RoboDK station: Bench V1 cell v7.rdk

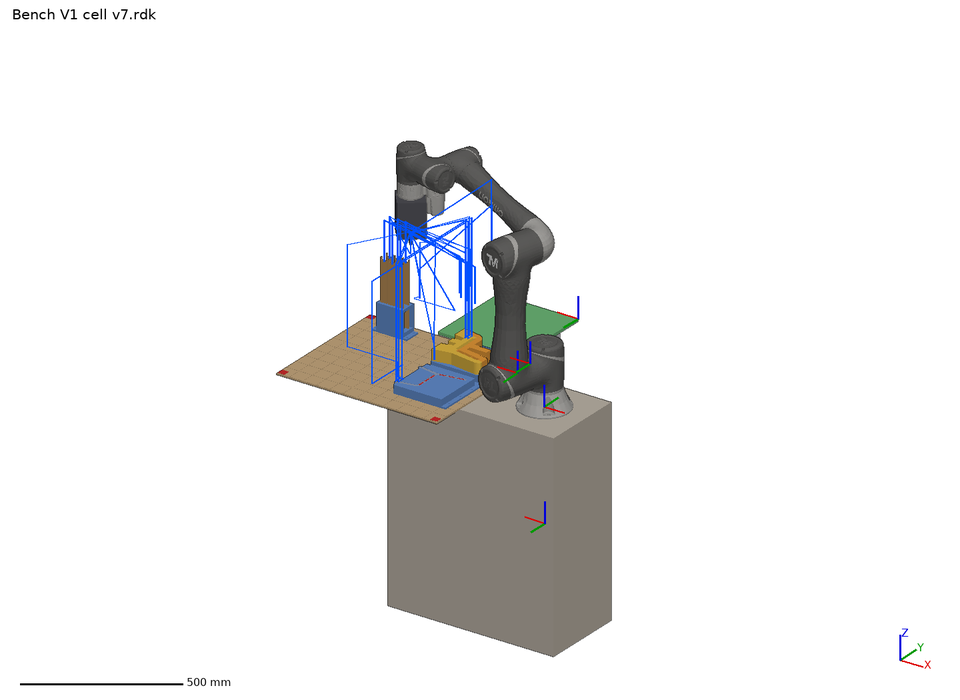
[picture v0: the station drawn from its stored meshes, robots at their saved joint values, targets as dots, program paths as lines]
Station Bench V1 cell v7 (saved by RoboDK 6.1.1). Poses are relative to the parent item; angles as X-Y-Z fixed-axis rotations.
  - frame Cell at (0, 0, 0) mm
    - frame Work plate at (-206.44, 152.99, -4.46) mm, rotated rx -0.03 ry -0.07 rz -179.98 deg
      - frame Ground base at (0, -67, 6) mm
        - object Table at (0, 0, 0) mm, size 620 x 310 x 744 mm
        - object Ground base plate at (0, 0, 0) mm, size 600 x 500 x 6 mm, geometry from ground_base_v7.stl
        - object Vision square 1 at (3, 3, 0) mm, size 25 x 25 x 0.5 mm, geometry from vision_square.stl
        - object Vision square 2 at (3, 472, 0) mm, size 25 x 25 x 0.5 mm, geometry from vision_square.stl
        - object Vision square 3 at (572, 3, 0) mm, size 25 x 25 x 0.5 mm, geometry from vision_square.stl
        - object Vision square 4 at (572, 472, 0) mm, size 25 x 25 x 0.5 mm, geometry from vision_square.stl
        - object Base A at (135, 122, 10) mm, rotated rx 0 ry 0 rz 90 deg, size 196 x 196 x 30 mm, geometry from base_a_v7.stl
        - object Base B at (135, 322, 10) mm, rotated rx 0 ry 0 rz -90 deg, size 196 x 196 x 30 mm, geometry from base_b_v7.stl
        - object Plank jig at (420, 30, 0) mm, size 132 x 60 x 100 mm, geometry from plank_rack_v7.stl
        - frame AMR at (60, -340, 0) mm
          - object AMR plate at (0, 0, 0) mm, size 300 x 320 x 10 mm
          - object AMR top module at (0, 0, 0) mm, size 220 x 240 x 363 mm
          - frame Omron LD-250 Base at (150, -40, -756) mm
            - robot AMR LD-250: 4 axes
                joint limits [-10000, -10000, -10, -3600] to [10000, 10000, 10, 3600]; home [0, 0, 0, 0]; saved at [0, 0, 0, 0]
        - object frame1 at (161.88, 119.28, 144.5) mm, size 174.7 x 141.9 x 10 mm, geometry from frame.stl
        - object frame2 at (161.88, 324.71, -95.5) mm, rotated rx 180 ry 0 rz 0 deg, size 174.7 x 141.9 x 10 mm, geometry from frame.stl
        - object piece A1 at (156.88, 119.28, 144.5) mm, rotated rx 90 ry 0 rz 90 deg, size 21.4 x 10 x 5 mm, geometry from interface_piece.stl
        - object piece B1 at (156.88, 324.71, 144.5) mm, rotated rx 90 ry 0 rz 90 deg, size 21.4 x 10 x 5 mm, geometry from interface_piece.stl
        - object plank1 at (435, 47.5, 128) mm, rotated rx 90 ry 0 rz 0 deg, size 25 x 250 x 5 mm, geometry from plank_body.stl
        - object piece A2 at (156.88, 89.3, 144.5) mm, rotated rx 90 ry 0 rz 90 deg, size 21.4 x 10 x 5 mm, geometry from interface_piece.stl
        - object piece B2 at (156.88, 354.7, 144.5) mm, rotated rx 90 ry 0 rz 90 deg, size 21.4 x 10 x 5 mm, geometry from interface_piece.stl
        - object plank2 at (465, 47.5, 128) mm, rotated rx 90 ry 0 rz 0 deg, size 25 x 250 x 5 mm, geometry from plank_body.stl
        - object piece A3 at (156.88, 149.27, 144.5) mm, rotated rx 90 ry 0 rz 90 deg, size 21.4 x 10 x 5 mm, geometry from interface_piece.stl
        - object piece B3 at (156.88, 294.73, 144.5) mm, rotated rx 90 ry 0 rz 90 deg, size 21.4 x 10 x 5 mm, geometry from interface_piece.stl
        - object plank3 at (495, 47.5, 128) mm, rotated rx 90 ry 0 rz 0 deg, size 25 x 250 x 5 mm, geometry from plank_body.stl
        - object piece A4 at (138.44, 171.24, 144.5) mm, rotated rx 90 ry 0 rz 170 deg, size 21.4 x 10 x 5 mm, geometry from interface_piece.stl
        - object piece B4 at (138.44, 272.76, 144.5) mm, rotated rx 90 ry 0 rz 10 deg, size 21.4 x 10 x 5 mm, geometry from interface_piece.stl
        - object plank4 at (435, 77.5, 128) mm, rotated rx 90 ry 0 rz 0 deg, size 25 x 250 x 5 mm, geometry from plank_body.stl
        - object piece A5 at (108.91, 176.45, 144.5) mm, rotated rx 90 ry 0 rz 170 deg, size 21.4 x 10 x 5 mm, geometry from interface_piece.stl
        - object piece B5 at (108.91, 267.55, 144.5) mm, rotated rx 90 ry 0 rz 10 deg, size 21.4 x 10 x 5 mm, geometry from interface_piece.stl
        - object plank5 at (465, 77.5, 128) mm, rotated rx 90 ry 0 rz 0 deg, size 25 x 250 x 5 mm, geometry from plank_body.stl
        - object piece A6 at (79.38, 181.66, 144.5) mm, rotated rx 90 ry 0 rz 170 deg, size 21.4 x 10 x 5 mm, geometry from interface_piece.stl
        - object piece B6 at (79.38, 262.34, 144.5) mm, rotated rx 90 ry 0 rz 10 deg, size 21.4 x 10 x 5 mm, geometry from interface_piece.stl
        - object plank6 at (495, 77.5, 128) mm, rotated rx 90 ry 0 rz 0 deg, size 25 x 250 x 5 mm, geometry from plank_body.stl
        - object Guide inner at (135, 122, 10) mm, rotated rx 0 ry 0 rz 90 deg, size 158.3 x 160 x 40 mm, geometry from guide_inner_v7.stl
        - object Guide outer at (135, 122, 10) mm, rotated rx 0 ry 0 rz 90 deg, size 177.7 x 180 x 40 mm, geometry from guide_outer_v7.stl
        - target Home (Cartesian target) at (295, 220, 380) mm, rotated rx 180 ry 0 rz 0 deg; joints [-14.089, 3.172, -81.623, -11.478, -90.01, 75.887] of Omron TM5-900
        - target plank3 pick travel (Cartesian target) at (495, 45, 380) mm, rotated rx 180 ry 0 rz -90 deg; joints [-23.734, -30.79, -38.937, -20.201, -89.998, 156.242] of Omron TM5-900
        - target plank3 pick approach (Cartesian target) at (495, 45, 278) mm, rotated rx 180 ry 0 rz -90 deg; joints [-23.733, -27.058, -59.189, -3.681, -89.998, 156.243] of Omron TM5-900
        - target plank3 pick (Cartesian target) at (495, 45, 238) mm, rotated rx 180 ry 0 rz -90 deg; joints [-23.733, -26.967, -64.904, 1.942, -89.998, 156.243] of Omron TM5-900
        - target plank3 pick out (Cartesian target) at (495, 45, 298) mm, rotated rx 180 ry 0 rz -90 deg; joints [-23.733, -27.342, -55.969, -6.617, -89.998, 156.243] of Omron TM5-900
        - target plank3 pick up (Cartesian target) at (495, 45, 380) mm, rotated rx 180 ry 0 rz -90 deg; joints [-23.734, -30.79, -38.937, -20.201, -89.998, 156.242] of Omron TM5-900
        - target plank3 place travel (Cartesian target) at (159.38, 149.27, 380) mm, rotated rx 180 ry 0 rz 0 deg; joints [-30.116, 20.707, -95.296, -15.34, -89.99, 59.86] of Omron TM5-900
        - target plank3 above guide (Cartesian target) at (159.38, 149.27, 329.5) mm, rotated rx 180 ry 0 rz 0 deg; joints [-30.114, 22.129, -103.368, -8.691, -89.99, 59.862] of Omron TM5-900
        - target plank3 place (Cartesian target) at (159.38, 149.27, 254.5) mm, rotated rx 180 ry 0 rz 0 deg; joints [-30.112, 22.789, -114.254, 1.536, -89.99, 59.864] of Omron TM5-900
        - target plank3 push approach (Cartesian target) at (159.38, 149.27, 289.5) mm, rotated rx 180 ry 0 rz 0 deg; joints [-30.113, 22.711, -109.326, -3.314, -89.99, 59.863] of Omron TM5-900
        - target plank3 push (Cartesian target) at (159.38, 149.27, 269.5) mm, rotated rx 180 ry 0 rz 0 deg; joints [-30.113, 22.808, -112.174, -0.563, -89.99, 59.863] of Omron TM5-900
        - target plank3 push out (Cartesian target) at (159.38, 149.27, 289.5) mm, rotated rx 180 ry 0 rz 0 deg; joints [-30.113, 22.711, -109.326, -3.314, -89.99, 59.863] of Omron TM5-900
        - target plank3 place up (Cartesian target) at (159.38, 149.27, 380) mm, rotated rx 180 ry 0 rz 0 deg; joints [-30.116, 20.707, -95.296, -15.34, -89.99, 59.86] of Omron TM5-900
        - target plank6 pick travel (Cartesian target) at (495, 75, 380) mm, rotated rx 180 ry 0 rz -90 deg; joints [-21.493, -29.466, -41.001, -19.462, -90.001, 158.482] of Omron TM5-900
        - target plank6 pick approach (Cartesian target) at (495, 75, 278) mm, rotated rx 180 ry 0 rz -90 deg; joints [-21.494, -26.016, -60.721, -3.192, -90.001, 158.482] of Omron TM5-900
        - target plank6 pick (Cartesian target) at (495, 75, 238) mm, rotated rx 180 ry 0 rz -90 deg; joints [-21.494, -25.975, -66.359, 2.406, -90.001, 158.482] of Omron TM5-900
        - target plank6 pick out (Cartesian target) at (495, 75, 298) mm, rotated rx 180 ry 0 rz -90 deg; joints [-21.494, -26.268, -57.554, -6.106, -90.001, 158.482] of Omron TM5-900
        - target plank6 pick up (Cartesian target) at (495, 75, 380) mm, rotated rx 180 ry 0 rz -90 deg; joints [-21.493, -29.466, -41.001, -19.462, -90.001, 158.482] of Omron TM5-900
        - target plank6 place travel (Cartesian target) at (79.82, 184.12, 380) mm, rotated rx 180 ry 0 rz 80 deg; joints [-32.257, 32.355, -101.249, -21.035, -89.987, -22.281] of Omron TM5-900
        - target plank6 above guide (Cartesian target) at (79.82, 184.12, 329.5) mm, rotated rx 180 ry 0 rz 80 deg; joints [-32.254, 34.514, -109.51, -14.934, -89.987, -22.278] of Omron TM5-900
        - target plank6 place (Cartesian target) at (79.82, 184.12, 254.5) mm, rotated rx 180 ry 0 rz 80 deg; joints [-32.25, 36.477, -120.901, -5.506, -89.987, -22.275] of Omron TM5-900
        - target plank6 push approach (Cartesian target) at (79.82, 184.12, 289.5) mm, rotated rx 180 ry 0 rz 80 deg; joints [-32.252, 35.762, -115.703, -9.988, -89.987, -22.276] of Omron TM5-900
        - target plank6 push (Cartesian target) at (79.82, 184.12, 269.5) mm, rotated rx 180 ry 0 rz 80 deg; joints [-32.251, 36.217, -118.697, -7.449, -89.987, -22.275] of Omron TM5-900
        - target plank6 push out (Cartesian target) at (79.82, 184.12, 289.5) mm, rotated rx 180 ry 0 rz 80 deg; joints [-32.252, 35.762, -115.703, -9.988, -89.987, -22.276] of Omron TM5-900
        - target plank6 place up (Cartesian target) at (79.82, 184.12, 380) mm, rotated rx 180 ry 0 rz 80 deg; joints [-32.257, 32.355, -101.249, -21.035, -89.987, -22.281] of Omron TM5-900
        - target plank2 pick travel (Cartesian target) at (465, 45, 380) mm, rotated rx 180 ry 0 rz -90 deg; joints [-24.747, -25.325, -47.241, -17.362, -89.997, 155.229] of Omron TM5-900
        - target plank2 pick approach (Cartesian target) at (465, 45, 278) mm, rotated rx 180 ry 0 rz -90 deg; joints [-24.747, -22.614, -65.589, -1.725, -89.997, 155.229] of Omron TM5-900
        - target plank2 pick (Cartesian target) at (465, 45, 238) mm, rotated rx 180 ry 0 rz -90 deg; joints [-24.746, -22.719, -71.021, 3.812, -89.997, 155.229] of Omron TM5-900
        - target plank2 pick out (Cartesian target) at (465, 45, 298) mm, rotated rx 180 ry 0 rz -90 deg; joints [-24.747, -22.777, -62.567, -4.584, -89.997, 155.229] of Omron TM5-900
        - target plank2 pick up (Cartesian target) at (465, 45, 380) mm, rotated rx 180 ry 0 rz -90 deg; joints [-24.747, -25.325, -47.241, -17.362, -89.997, 155.229] of Omron TM5-900
        - target plank2 place travel (Cartesian target) at (159.38, 89.3, 380) mm, rotated rx 180 ry 0 rz 0 deg; joints [-38.038, 18.536, -93.909, -14.558, -89.98, 51.938] of Omron TM5-900
        - target plank2 above guide (Cartesian target) at (159.38, 89.3, 329.5) mm, rotated rx 180 ry 0 rz 0 deg; joints [-38.035, 19.858, -101.95, -7.839, -89.98, 51.941] of Omron TM5-900
        - target plank2 place (Cartesian target) at (159.38, 89.3, 254.5) mm, rotated rx 180 ry 0 rz 0 deg; joints [-38.031, 20.348, -112.746, 2.466, -89.98, 51.945] of Omron TM5-900
        - target plank2 push approach (Cartesian target) at (159.38, 89.3, 289.5) mm, rotated rx 180 ry 0 rz 0 deg; joints [-38.033, 20.351, -107.867, -2.415, -89.98, 51.943] of Omron TM5-900
        - target plank2 push (Cartesian target) at (159.38, 89.3, 269.5) mm, rotated rx 180 ry 0 rz 0 deg; joints [-38.032, 20.402, -110.688, 0.355, -89.98, 51.944] of Omron TM5-900
        - target plank2 push out (Cartesian target) at (159.38, 89.3, 289.5) mm, rotated rx 180 ry 0 rz 0 deg; joints [-38.033, 20.351, -107.867, -2.415, -89.98, 51.943] of Omron TM5-900
        - target plank2 place up (Cartesian target) at (159.38, 89.3, 380) mm, rotated rx 180 ry 0 rz 0 deg; joints [-38.038, 18.536, -93.909, -14.558, -89.98, 51.938] of Omron TM5-900
        - target plank5 pick travel (Cartesian target) at (465, 75, 380) mm, rotated rx 180 ry 0 rz -90 deg; joints [-22.426, -24.114, -49.008, -16.806, -90, 157.55] of Omron TM5-900
        - target plank5 pick approach (Cartesian target) at (465, 75, 278) mm, rotated rx 180 ry 0 rz -90 deg; joints [-22.426, -21.584, -67.026, -1.319, -90, 157.55] of Omron TM5-900
        - target plank5 pick (Cartesian target) at (465, 75, 238) mm, rotated rx 180 ry 0 rz -90 deg; joints [-22.426, -21.727, -72.407, 4.206, -90, 157.55] of Omron TM5-900
        - target plank5 pick out (Cartesian target) at (465, 75, 298) mm, rotated rx 180 ry 0 rz -90 deg; joints [-22.426, -21.724, -64.039, -4.165, -90, 157.55] of Omron TM5-900
        - target plank5 pick up (Cartesian target) at (465, 75, 380) mm, rotated rx 180 ry 0 rz -90 deg; joints [-22.426, -24.114, -49.008, -16.806, -90, 157.55] of Omron TM5-900
        - target plank5 place travel (Cartesian target) at (109.34, 178.91, 380) mm, rotated rx 180 ry 0 rz 80 deg; joints [-30.015, 28.172, -99.401, -18.7, -89.99, -20.039] of Omron TM5-900
        - target plank5 above guide (Cartesian target) at (109.34, 178.91, 329.5) mm, rotated rx 180 ry 0 rz 80 deg; joints [-30.014, 30.03, -107.592, -12.366, -89.99, -20.038] of Omron TM5-900
        - target plank5 place (Cartesian target) at (109.34, 178.91, 254.5) mm, rotated rx 180 ry 0 rz 80 deg; joints [-30.011, 31.445, -118.805, -2.57, -89.99, -20.035] of Omron TM5-900
        - target plank5 push approach (Cartesian target) at (109.34, 178.91, 289.5) mm, rotated rx 180 ry 0 rz 80 deg; joints [-30.012, 31.001, -113.703, -7.227, -89.99, -20.036] of Omron TM5-900
        - target plank5 push (Cartesian target) at (109.34, 178.91, 269.5) mm, rotated rx 180 ry 0 rz 80 deg; joints [-30.012, 31.304, -116.645, -4.588, -89.99, -20.036] of Omron TM5-900
        - target plank5 push out (Cartesian target) at (109.34, 178.91, 289.5) mm, rotated rx 180 ry 0 rz 80 deg; joints [-30.012, 31.001, -113.703, -7.227, -89.99, -20.036] of Omron TM5-900
        - target plank5 place up (Cartesian target) at (109.34, 178.91, 380) mm, rotated rx 180 ry 0 rz 80 deg; joints [-30.015, 28.172, -99.401, -18.7, -89.99, -20.039] of Omron TM5-900
        - target plank1 pick travel (Cartesian target) at (435, 45, 380) mm, rotated rx 180 ry 0 rz -90 deg; joints [-25.849, -20.444, -54.192, -15.292, -89.995, 154.127] of Omron TM5-900
        - target plank1 pick approach (Cartesian target) at (435, 45, 278) mm, rotated rx 180 ry 0 rz -90 deg; joints [-25.848, -18.383, -71.372, -0.174, -89.995, 154.128] of Omron TM5-900
        - target plank1 pick (Cartesian target) at (435, 45, 238) mm, rotated rx 180 ry 0 rz -90 deg; joints [-25.848, -18.633, -76.622, 5.327, -89.995, 154.128] of Omron TM5-900
        - target plank1 pick out (Cartesian target) at (435, 45, 298) mm, rotated rx 180 ry 0 rz -90 deg; joints [-25.848, -18.461, -68.478, -2.99, -89.995, 154.128] of Omron TM5-900
        - target plank1 pick up (Cartesian target) at (435, 45, 380) mm, rotated rx 180 ry 0 rz -90 deg; joints [-25.849, -20.444, -54.192, -15.292, -89.995, 154.127] of Omron TM5-900
        - target plank1 place travel (Cartesian target) at (159.38, 119.28, 380) mm, rotated rx 180 ry 0 rz 0 deg; joints [-34.216, 19.771, -94.709, -14.993, -89.985, 55.76] of Omron TM5-900
        - target plank1 above guide (Cartesian target) at (159.38, 119.28, 329.5) mm, rotated rx 180 ry 0 rz 0 deg; joints [-34.214, 21.149, -102.767, -8.312, -89.985, 55.762] of Omron TM5-900
        - target plank1 place (Cartesian target) at (159.38, 119.28, 254.5) mm, rotated rx 180 ry 0 rz 0 deg; joints [-34.211, 21.733, -113.614, 1.951, -89.985, 55.765] of Omron TM5-900
        - target plank1 push approach (Cartesian target) at (159.38, 119.28, 289.5) mm, rotated rx 180 ry 0 rz 0 deg; joints [-34.212, 21.691, -108.707, -2.914, -89.985, 55.764] of Omron TM5-900
        - target plank1 push (Cartesian target) at (159.38, 119.28, 269.5) mm, rotated rx 180 ry 0 rz 0 deg; joints [-34.211, 21.767, -111.543, -0.154, -89.985, 55.764] of Omron TM5-900
        - target plank1 push out (Cartesian target) at (159.38, 119.28, 289.5) mm, rotated rx 180 ry 0 rz 0 deg; joints [-34.212, 21.691, -108.707, -2.914, -89.985, 55.764] of Omron TM5-900
        - target plank1 place up (Cartesian target) at (159.38, 119.28, 380) mm, rotated rx 180 ry 0 rz 0 deg; joints [-34.216, 19.771, -94.709, -14.993, -89.985, 55.76] of Omron TM5-900
        - target plank4 pick travel (Cartesian target) at (435, 75, 380) mm, rotated rx 180 ry 0 rz -90 deg; joints [-23.442, -19.281, -55.785, -14.863, -89.998, 156.534] of Omron TM5-900
        - target plank4 pick approach (Cartesian target) at (435, 75, 278) mm, rotated rx 180 ry 0 rz -90 deg; joints [-23.441, -17.346, -72.742, 0.16, -89.998, 156.535] of Omron TM5-900
        - target plank4 pick (Cartesian target) at (435, 75, 238) mm, rotated rx 180 ry 0 rz -90 deg; joints [-23.441, -17.626, -77.959, 5.657, -89.998, 156.535] of Omron TM5-900
        - target plank4 pick out (Cartesian target) at (435, 75, 298) mm, rotated rx 180 ry 0 rz -90 deg; joints [-23.441, -17.407, -69.873, -2.648, -89.998, 156.534] of Omron TM5-900
        - target plank4 pick up (Cartesian target) at (435, 75, 380) mm, rotated rx 180 ry 0 rz -90 deg; joints [-23.442, -19.281, -55.785, -14.863, -89.998, 156.534] of Omron TM5-900
        - target plank4 place travel (Cartesian target) at (138.87, 173.7, 380) mm, rotated rx 180 ry 0 rz 80 deg; joints [-28.195, 24.029, -97.25, -16.707, -89.992, -18.219] of Omron TM5-900
        - target plank4 above guide (Cartesian target) at (138.87, 173.7, 329.5) mm, rotated rx 180 ry 0 rz 80 deg; joints [-28.193, 25.628, -105.373, -10.184, -89.992, -18.218] of Omron TM5-900
        - target plank4 place (Cartesian target) at (138.87, 173.7, 254.5) mm, rotated rx 180 ry 0 rz 80 deg; joints [-28.192, 26.59, -116.403, -0.116, -89.992, -18.216] of Omron TM5-900
        - target plank4 push approach (Cartesian target) at (138.87, 173.7, 289.5) mm, rotated rx 180 ry 0 rz 80 deg; joints [-28.193, 26.366, -111.398, -4.897, -89.992, -18.217] of Omron TM5-900
        - target plank4 push (Cartesian target) at (138.87, 173.7, 269.5) mm, rotated rx 180 ry 0 rz 80 deg; joints [-28.192, 26.545, -114.287, -2.187, -89.992, -18.216] of Omron TM5-900
        - target plank4 push out (Cartesian target) at (138.87, 173.7, 289.5) mm, rotated rx 180 ry 0 rz 80 deg; joints [-28.193, 26.366, -111.398, -4.897, -89.992, -18.217] of Omron TM5-900
        - target plank4 place up (Cartesian target) at (138.87, 173.7, 380) mm, rotated rx 180 ry 0 rz 80 deg; joints [-28.195, 24.029, -97.25, -16.707, -89.992, -18.219] of Omron TM5-900
        - target guide A-B pick out low (Cartesian target) at (205, 25, 50) mm, rotated rx 0 ry -90 rz -90 deg; joints [-60.041, -46.665, -86.504, -46.801, -60.065, -90.051] of Omron TM5-900
        - target guide A-B pick out (Cartesian target) at (205, 25, 450) mm, rotated rx 0 ry -90 rz -90 deg; joints [-60.07, -28.06, -57.103, -94.806, -60.094, -90.051] of Omron TM5-900
        - target guide A-B via (Cartesian target) at (295, 220, 450) mm, rotated rx 0 ry -90 rz -90 deg; joints [-41.029, -19.995, -68.597, -91.367, -41.053, -90.035] of Omron TM5-900
        - target guide A-B pick (Cartesian target) at (205, 50, 50) mm, rotated rx 0 ry -90 rz -90 deg; joints [-58.833, -44.847, -90.216, -44.905, -58.857, -90.05] of Omron TM5-900
        - target guide A-B lift (Cartesian target) at (205, 50, 70) mm, rotated rx 0 ry -90 rz -90 deg; joints [-58.834, -42.987, -90.07, -46.911, -58.858, -90.05] of Omron TM5-900
        - target guide A-B up (Cartesian target) at (205, 50, 450) mm, rotated rx 0 ry -90 rz -90 deg; joints [-58.862, -25.121, -61.421, -93.427, -58.886, -90.05] of Omron TM5-900
        - target guide A-B across (Cartesian target) at (205, 394, 450) mm, rotated rx 0 ry -90 rz -90 deg; joints [-30.469, 0.804, -93.022, -87.729, -30.493, -90.021] of Omron TM5-900
        - target guide A-B place (Cartesian target) at (205, 394, 50) mm, rotated rx 0 ry 90 rz -90 deg; joints [35.876, -45.178, -89.623, -45.245, -144.148, -269.896] of Omron TM5-900
        - target guide A-B over place (Cartesian target) at (205, 394, 450) mm, rotated rx 0 ry 90 rz -90 deg; joints [35.917, -25.629, -60.744, -93.673, -144.107, -269.896] of Omron TM5-900
        - target guide A-B place approach (Cartesian target) at (205, 394, 90) mm, rotated rx 0 ry 90 rz -90 deg; joints [35.88, -41.547, -89.201, -49.298, -144.144, -269.896] of Omron TM5-900
        - target guide A-B place out (Cartesian target) at (205, 419, 50) mm, rotated rx 0 ry 90 rz -90 deg; joints [37.771, -47.012, -85.878, -47.153, -142.253, -269.899] of Omron TM5-900
        - target guide A-B place out up (Cartesian target) at (205, 419, 450) mm, rotated rx 0 ry 90 rz -90 deg; joints [37.811, -28.6, -56.357, -95.087, -142.213, -269.899] of Omron TM5-900
        - target sub pick (Cartesian target) at (231.7, 182.8, 22) mm, rotated rx -120 ry 0 rz 99.93 deg; joints [-10.147, -38.104, -86.099, -24.148, -107.32, -10.354] of Omron TM5-900
        - target sub pick approach (Cartesian target) at (231.7, 182.8, 62) mm, rotated rx -120 ry 0 rz 99.93 deg; joints [-10.147, -35.261, -84.458, -28.633, -107.32, -10.354] of Omron TM5-900
        - target sub via (Cartesian target) at (295, 220, 450) mm, rotated rx -120 ry 0 rz 99.93 deg; joints [-10.147, -38.104, -86.099, -24.148, -107.32, -10.354] of Omron TM5-900
        - target sub to middle (joint target) at (200, 222, 450) mm, rotated rx -120 ry 0 rz 99.93 deg; joints [-7.117, -26.573, -41.835, -80.397, -104.734, -8.711] of Omron TM5-900
        - target sub place (Cartesian target) at (231.7, 261.2, 267) mm, rotated rx 60 ry 0 rz -99.93 deg; joints [-10.443, -53.16, -62.534, -94.237, -90.461, -179.717] of Omron TM5-900
        - target sub above guide (Cartesian target) at (231.7, 261.2, 342) mm, rotated rx 60 ry 0 rz -99.93 deg; joints [-10.441, -48.865, -59.308, -101.758, -90.46, -179.718] of Omron TM5-900
        - target sub flipped high (Cartesian target) at (231.7, 261.2, 450) mm, rotated rx 60 ry 0 rz -99.93 deg; joints [-10.439, -45.209, -50.407, -114.316, -90.457, -179.719] of Omron TM5-900
        - target sub flipped (Cartesian target) at (231.7, 261.2, 387) mm, rotated rx 60 ry 0 rz -99.93 deg; joints [-10.44, -46.936, -56.271, -106.724, -90.459, -179.718] of Omron TM5-900
        - target sub place out (Cartesian target) at (253.03, 257.47, 254.5) mm, rotated rx 60 ry 0 rz -99.93 deg; joints [-10.426, -57.015, -56.959, -95.957, -90.446, -179.726] of Omron TM5-900
        - target sub clear (Cartesian target) at (103.03, 257.47, 254.5) mm, rotated rx 60 ry 0 rz -99.93 deg; joints [-13.356, -39, -91.524, -79.451, -92.985, -178.262] of Omron TM5-900
        - target sub back to middle (Cartesian target) at (295, 220, 450) mm, rotated rx 60 ry 0 rz -99.93 deg; joints [-12.723, -59.734, -23.858, -126.368, -92.436, -178.579] of Omron TM5-900
        - target outer pick out low (Cartesian target) at (210, 419, 50) mm, rotated rx 0 ry 90 rz -90 deg; joints [37.488, -47.342, -85.204, -47.498, -142.537, 90.102] of Omron TM5-900
        - target outer pick out (Cartesian target) at (210, 419, 450) mm, rotated rx 0 ry 90 rz -90 deg; joints [37.528, -29.139, -55.545, -95.361, -142.497, 90.102] of Omron TM5-900
        - target outer via (Cartesian target) at (295, 220, 450) mm, rotated rx 0 ry 90 rz -90 deg; joints [16.365, -20.051, -68.557, -91.488, -163.659, 90.158] of Omron TM5-900
        - target outer pick (Cartesian target) at (210, 394, 50) mm, rotated rx 0 ry 90 rz -90 deg; joints [35.596, -45.506, -88.951, -45.589, -144.428, 90.104] of Omron TM5-900
        - target outer out 1 (Cartesian target) at (218, 394, 50) mm, rotated rx 0 ry 90 rz -90 deg; joints [35.156, -46.041, -87.857, -46.149, -144.868, 90.105] of Omron TM5-900
        - target outer out 2 (Cartesian target) at (218, 394, 100) mm, rotated rx 0 ry 90 rz -90 deg; joints [35.161, -41.619, -87.247, -51.181, -144.863, 90.105] of Omron TM5-900
        - target outer out 3 (Cartesian target) at (408, 394, 100) mm, rotated rx 0 ry 90 rz -90 deg; joints [26.881, -59.522, -52.568, -67.97, -153.143, 90.12] of Omron TM5-900
        - target outer up (Cartesian target) at (408, 394, 450) mm, rotated rx 0 ry 90 rz -90 deg; joints [26.906, -53.115, -44.921, 97.977, 153.118, -89.88] of Omron TM5-900
        - target outer across (Cartesian target) at (210, 50, 450) mm, rotated rx 0 ry 90 rz -90 deg; joints [-2.472, 0.124, -92.361, -87.144, 177.504, 89.448] of Omron TM5-900
        - target outer place (Cartesian target) at (210, 50, 50) mm, rotated rx 0 ry -90 rz -90 deg; joints [-58.421, -45.176, -89.544, -45.249, -58.445, -90.05] of Omron TM5-900
        - target outer over place (Cartesian target) at (210, 50, 450) mm, rotated rx 0 ry -90 rz -90 deg; joints [-58.45, -25.651, -60.652, -93.665, -58.474, -90.05] of Omron TM5-900
        - target outer place approach (Cartesian target) at (210, 50, 90) mm, rotated rx 0 ry -90 rz -90 deg; joints [-58.424, -41.548, -89.121, -49.299, -58.448, -90.05] of Omron TM5-900
        - target outer place out (Cartesian target) at (210, 25, 50) mm, rotated rx 0 ry -90 rz -90 deg; joints [-59.637, -46.994, -85.83, -47.145, -59.661, -90.051] of Omron TM5-900
        - target outer place out up (Cartesian target) at (210, 25, 450) mm, rotated rx 0 ry -90 rz -90 deg; joints [-59.666, -28.597, -56.299, -95.073, -59.69, -90.051] of Omron TM5-900
        - target inner pick out low (Cartesian target) at (200, 419, 50) mm, rotated rx 0 ry 90 rz -90 deg; joints [38.058, -46.687, -86.544, -46.813, -141.966, 90.101] of Omron TM5-900
        - target inner pick out (Cartesian target) at (200, 419, 450) mm, rotated rx 0 ry 90 rz -90 deg; joints [38.099, -28.07, -57.151, -94.822, -141.925, 90.101] of Omron TM5-900
        - target inner via (Cartesian target) at (295, 220, 450) mm, rotated rx 0 ry 90 rz -90 deg; joints [16.365, -20.051, -68.557, -91.488, -163.659, 90.158] of Omron TM5-900
        - target inner pick (Cartesian target) at (200, 394, 50) mm, rotated rx 0 ry 90 rz -90 deg; joints [36.16, -44.853, -90.288, -44.905, -143.864, 90.103] of Omron TM5-900
        - target inner out 1 (Cartesian target) at (198.61, 401.88, 50) mm, rotated rx 0 ry 90 rz -90 deg; joints [36.849, -45.33, -89.314, -45.401, -143.175, 90.102] of Omron TM5-900
        - target inner out 2 (Cartesian target) at (198.61, 401.88, 100) mm, rotated rx 0 ry 90 rz -90 deg; joints [36.854, -40.85, -88.704, -50.491, -143.17, 90.102] of Omron TM5-900
        - target inner out 3 (Cartesian target) at (198.61, 561.88, 100) mm, rotated rx 0 ry 90 rz -90 deg; joints [47.16, -56.068, -59.404, -64.565, -132.865, 90.091] of Omron TM5-900
        - target inner up (Cartesian target) at (198.61, 561.88, 450) mm, rotated rx 0 ry 90 rz -90 deg; joints [47.192, -54.867, -11.337, -113.833, -132.832, 90.091] of Omron TM5-900
        - target inner across (Cartesian target) at (200, 50, 450) mm, rotated rx 0 ry 90 rz -90 deg; joints [-2.534, -119.323, 115.434, 4.493, -177.442, 269.463] of Omron TM5-900
        - target inner place (Cartesian target) at (200, 50, 50) mm, rotated rx 0 ry -90 rz -90 deg; joints [-59.248, -44.523, -90.88, -44.566, -59.272, 269.95] of Omron TM5-900
        - target inner over place (Cartesian target) at (200, 50, 450) mm, rotated rx 0 ry -90 rz -90 deg; joints [-59.278, -24.598, -62.174, -93.196, -59.302, 269.95] of Omron TM5-900
        - target inner place approach (Cartesian target) at (200, 50, 90) mm, rotated rx 0 ry -90 rz -90 deg; joints [-59.251, -40.85, -90.457, -48.662, -59.275, 269.95] of Omron TM5-900
        - target inner place out (Cartesian target) at (200, 25, 50) mm, rotated rx 0 ry -90 rz -90 deg; joints [-60.449, -46.339, -87.169, -46.461, -60.473, 269.949] of Omron TM5-900
        - target inner place out up (Cartesian target) at (200, 25, 450) mm, rotated rx 0 ry -90 rz -90 deg; joints [-60.478, -27.532, -57.891, -94.547, -60.502, 269.949] of Omron TM5-900
        - target bench pick out low (Cartesian target) at (231.7, 261.2, 287) mm, rotated rx 180 ry 0 rz -99.93 deg; joints [-10.732, 12.862, -102.959, 0.168, -90.014, 179.17] of Omron TM5-900
        - target bench pick out (Cartesian target) at (231.7, 261.2, 322) mm, rotated rx 180 ry 0 rz -99.93 deg; joints [-10.731, 12.674, -97.931, -4.674, -90.014, 179.171] of Omron TM5-900
        - target bench via (Cartesian target) at (295, 220, 450) mm, rotated rx 180 ry 0 rz -99.93 deg; joints [-14.088, 0.421, -68.77, -21.58, -90.01, 175.814] of Omron TM5-900
        - target bench pick (Cartesian target) at (231.7, 261.2, 262) mm, rotated rx 180 ry 0 rz -99.93 deg; joints [-10.733, 12.746, -106.358, 3.682, -90.014, 179.169] of Omron TM5-900
        - target bench lift (Cartesian target) at (231.7, 261.2, 362) mm, rotated rx 180 ry 0 rz -99.93 deg; joints [-10.729, 11.983, -91.768, -10.144, -90.014, 179.173] of Omron TM5-900
        - target bench over AMR (Cartesian target) at (305.7, -228.8, 362) mm, rotated rx 180 ry 0 rz -99.93 deg; joints [-51.593, -22.33, -54.157, -13.451, -89.965, 138.309] of Omron TM5-900
        - target bench down (Cartesian target) at (305.7, -228.8, 243) mm, rotated rx 180 ry 0 rz -99.93 deg; joints [-51.587, -20.844, -72.93, 3.837, -89.965, 138.315] of Omron TM5-900
        - target bench place out (Cartesian target) at (305.7, -228.8, 283) mm, rotated rx 180 ry 0 rz -99.93 deg; joints [-51.589, -20.738, -67.497, -1.703, -89.965, 138.313] of Omron TM5-900
        - target bench place out up (Cartesian target) at (305.7, -228.8, 450) mm, rotated rx 180 ry 0 rz -99.93 deg; joints [-51.598, -28.705, -31.441, -29.791, -89.965, 138.304] of Omron TM5-900
        - target back to middle (Cartesian target) at (295, 220, 450) mm, rotated rx -180 ry 0 rz -99.93 deg; joints [-14.088, 0.421, -68.769, -21.58, -90.01, 175.814] of Omron TM5-900
    - frame Omron TM5-900 Base at (0, 0, 0) mm
      - robot Omron TM5-900: 6 axes, payload 4 kg, reach 900 mm, repeatability 0.05 mm, weight 22.6 kg
          modified DH rows (alpha deg, a mm, theta deg, d mm): 0, 0, 0, 145.2; 90, 0, 90, 0; 0, 429, 0, 0; 0, 411, -90, 122.3; -90, 0, 0, 106.5; 90, 0, 180, 114.15
          joint limits [-270, -180, -155, -180, -180, -270] to [270, 180, 155, 180, 180, 270]; home [0, 0, 90, -90, 90, 0]; saved at [-14.089, 2.021, -75.497, -16.453, -90.01, 125.85]
        - tool EGP, TCP at (0, 0, 160) mm, size 94 x 90 x 160 mm
  - program AssembleBench (317 instructions, listed below)
  - Python program Deliver (AMR) (listed below)
  - Python program Assemble and deliver (listed below)
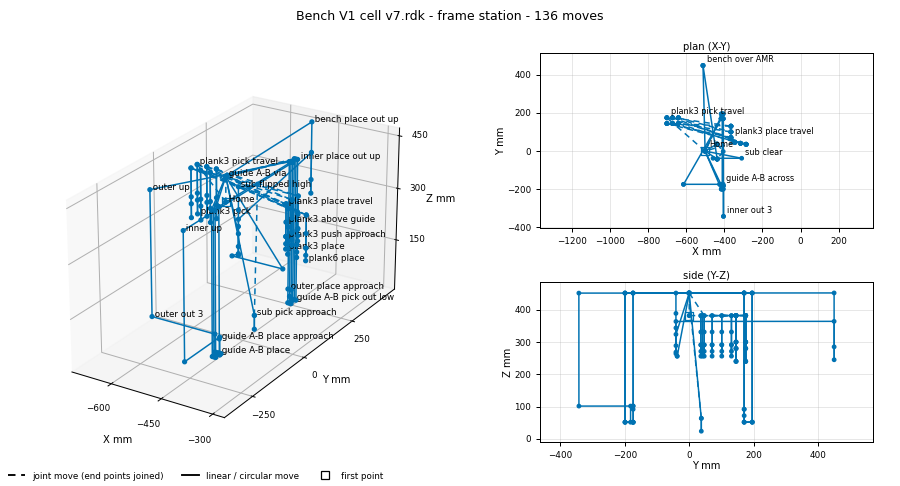
[picture p0: tool path of Bench V1 cell v7.rdk in frame station, 136 of 136 moves have a stored position in this frame; points joined in program order, loops and branches not executed]

--- program AssembleBench (robot Omron TM5-900) ---
  Simulation: parts to start
  Set Ref.: Ground base
  Set Tool: EGP
  Smooth(0)
  Set speed (100.0 mm/s)
  MoveJ (Home)
  MoveJ (plank3 pick travel)
  MoveL (plank3 pick approach)
  Set speed (20.0 mm/s)
  MoveL (plank3 pick)
  Set IO_0=1
  Pause 500 ms
  Simulation: attach plank3
  MoveL (plank3 pick out)
  Set speed (100.0 mm/s)
  MoveL (plank3 pick up)
  MoveJ (plank3 place travel)
  MoveL (plank3 above guide)
  Set speed (20.0 mm/s)
  MoveL (plank3 place)
  Set IO_0=0
  Pause 500 ms
  Simulation: release plank3
  MoveL (plank3 push approach)
  Set IO_0=1
  Pause 300 ms
  MoveL (plank3 push)
  MoveL (plank3 push out)
  Set IO_0=0
  Pause 300 ms
  Set speed (100.0 mm/s)
  MoveL (plank3 place up)
  MoveJ (plank6 pick travel)
  MoveL (plank6 pick approach)
  Set speed (20.0 mm/s)
  MoveL (plank6 pick)
  Set IO_0=1
  Pause 500 ms
  Simulation: attach plank6
  MoveL (plank6 pick out)
  Set speed (100.0 mm/s)
  MoveL (plank6 pick up)
  MoveJ (plank6 place travel)
  MoveL (plank6 above guide)
  Set speed (20.0 mm/s)
  MoveL (plank6 place)
  Set IO_0=0
  Pause 500 ms
  Simulation: release plank6
  MoveL (plank6 push approach)
  Set IO_0=1
  Pause 300 ms
  MoveL (plank6 push)
  MoveL (plank6 push out)
  Set IO_0=0
  Pause 300 ms
  Set speed (100.0 mm/s)
  MoveL (plank6 place up)
  MoveJ (plank2 pick travel)
  MoveL (plank2 pick approach)
  Set speed (20.0 mm/s)
  MoveL (plank2 pick)
  Set IO_0=1
  Pause 500 ms
  Simulation: attach plank2
  MoveL (plank2 pick out)
  Set speed (100.0 mm/s)
  MoveL (plank2 pick up)
  MoveJ (plank2 place travel)
  MoveL (plank2 above guide)
  Set speed (20.0 mm/s)
  MoveL (plank2 place)
  Set IO_0=0
  Pause 500 ms
  Simulation: release plank2
  MoveL (plank2 push approach)
  Set IO_0=1
  Pause 300 ms
  MoveL (plank2 push)
  MoveL (plank2 push out)
  Set IO_0=0
  Pause 300 ms
  Set speed (100.0 mm/s)
  MoveL (plank2 place up)
  MoveJ (plank5 pick travel)
  MoveL (plank5 pick approach)
  Set speed (20.0 mm/s)
  MoveL (plank5 pick)
  Set IO_0=1
  Pause 500 ms
  Simulation: attach plank5
  MoveL (plank5 pick out)
  Set speed (100.0 mm/s)
  MoveL (plank5 pick up)
  MoveJ (plank5 place travel)
  MoveL (plank5 above guide)
  Set speed (20.0 mm/s)
  MoveL (plank5 place)
  Set IO_0=0
  Pause 500 ms
  Simulation: release plank5
  MoveL (plank5 push approach)
  Set IO_0=1
  Pause 300 ms
  MoveL (plank5 push)
  MoveL (plank5 push out)
  Set IO_0=0
  Pause 300 ms
  Set speed (100.0 mm/s)
  MoveL (plank5 place up)
  MoveJ (plank1 pick travel)
  MoveL (plank1 pick approach)
  Set speed (20.0 mm/s)
  MoveL (plank1 pick)
  Set IO_0=1
  Pause 500 ms
  Simulation: attach plank1
  MoveL (plank1 pick out)
  Set speed (100.0 mm/s)
  MoveL (plank1 pick up)
  MoveJ (plank1 place travel)
  MoveL (plank1 above guide)
  Set speed (20.0 mm/s)
  MoveL (plank1 place)
  Set IO_0=0
  Pause 500 ms
  Simulation: release plank1
  MoveL (plank1 push approach)
  Set IO_0=1
  Pause 300 ms
  MoveL (plank1 push)
  MoveL (plank1 push out)
  Set IO_0=0
  Pause 300 ms
  Set speed (100.0 mm/s)
  MoveL (plank1 place up)
  MoveJ (plank4 pick travel)
  MoveL (plank4 pick approach)
  Set speed (20.0 mm/s)
  MoveL (plank4 pick)
  Set IO_0=1
  Pause 500 ms
  Simulation: attach plank4
  MoveL (plank4 pick out)
  Set speed (100.0 mm/s)
  MoveL (plank4 pick up)
  MoveJ (plank4 place travel)
  MoveL (plank4 above guide)
  Set speed (20.0 mm/s)
  MoveL (plank4 place)
  Set IO_0=0
  Pause 500 ms
  Simulation: release plank4
  MoveL (plank4 push approach)
  Set IO_0=1
  Pause 300 ms
  MoveL (plank4 push)
  MoveL (plank4 push out)
  Set IO_0=0
  Pause 300 ms
  Set speed (100.0 mm/s)
  MoveL (plank4 place up)
  MoveJ (guide A-B via)
  MoveL (guide A-B pick out)
  MoveL (guide A-B pick out low)
  Set speed (20.0 mm/s)
  Set IO_0=1
  Pause 300 ms
  MoveL (guide A-B pick)
  Set IO_0=0
  Pause 500 ms
  Simulation: attach Guide inner
  Simulation: attach Guide outer
  MoveL (guide A-B lift)
  Set speed (100.0 mm/s)
  MoveL (guide A-B up)
  MoveL (guide A-B across)
  MoveJ (guide A-B over place)
  MoveL (guide A-B place approach)
  Set speed (20.0 mm/s)
  MoveL (guide A-B place)
  Set IO_0=1
  Pause 500 ms
  Simulation: release guide A-B
  MoveL (guide A-B place out)
  Set speed (100.0 mm/s)
  MoveL (guide A-B place out up)
  MoveJ (sub via)
  MoveL (sub pick approach)
  Set speed (20.0 mm/s)
  MoveL (sub pick)
  Set IO_0=1
  Pause 500 ms
  Simulation: attach frame1
  Simulation: attach plank1
  Simulation: attach plank2
  Simulation: attach plank3
  Simulation: attach plank4
  Simulation: attach plank5
  Simulation: attach plank6
  Simulation: attach piece A1
  Simulation: attach piece A2
  Simulation: attach piece A3
  Simulation: attach piece A4
  Simulation: attach piece A5
  Simulation: attach piece A6
  MoveL (sub pick approach)
  Set speed (100.0 mm/s)
  MoveJ (sub to middle)
  MoveJ (sub flipped high)
  MoveL (sub flipped)
  MoveL (sub above guide)
  Set speed (20.0 mm/s)
  MoveL (sub place)
  Set IO_0=0
  Pause 500 ms
  Simulation: release frame 1 with the planks
  MoveL (sub place out)
  MoveL (sub clear)
  MoveL (sub back to middle)
  Set speed (100.0 mm/s)
  MoveJ (outer via)
  MoveL (outer pick out)
  MoveL (outer pick out low)
  Set speed (20.0 mm/s)
  Set IO_0=1
  Pause 300 ms
  MoveL (outer pick)
  Set IO_0=0
  Pause 500 ms
  Simulation: attach Guide outer
  Set speed (20.0 mm/s)
  MoveL (outer out 1)
  MoveL (outer out 2)
  MoveL (outer out 3)
  Set speed (100.0 mm/s)
  MoveL (outer up)
  MoveL (outer across)
  MoveJ (outer over place)
  MoveL (outer place approach)
  Set speed (20.0 mm/s)
  MoveL (outer place)
  Set IO_0=1
  Pause 500 ms
  Simulation: release outer
  MoveL (outer place out)
  Set speed (100.0 mm/s)
  MoveL (outer place out up)
  MoveJ (inner via)
  MoveL (inner pick out)
  MoveL (inner pick out low)
  Set speed (20.0 mm/s)
  Set IO_0=1
  Pause 300 ms
  MoveL (inner pick)
  Set IO_0=0
  Pause 500 ms
  Simulation: attach Guide inner
  Set speed (20.0 mm/s)
  MoveL (inner out 1)
  MoveL (inner out 2)
  MoveL (inner out 3)
  Set speed (100.0 mm/s)
  MoveL (inner up)
  MoveL (inner across)
  MoveJ (inner over place)
  MoveL (inner place approach)
  Set speed (20.0 mm/s)
  MoveL (inner place)
  Set IO_0=1
  Pause 500 ms
  Simulation: release inner
  MoveL (inner place out)
  Set speed (100.0 mm/s)
  MoveL (inner place out up)
  MoveJ (bench via)
  MoveL (bench pick out)
  MoveL (bench pick out low)
  Set speed (20.0 mm/s)
  Set IO_0=0
  Pause 300 ms
  MoveL (bench pick)
  Set IO_0=1
  Pause 500 ms
  Simulation: attach frame1
  Simulation: attach frame2
  Simulation: attach plank1
  Simulation: attach plank2
  Simulation: attach plank3
  Simulation: attach plank4
  Simulation: attach plank5
  Simulation: attach plank6
  Simulation: attach piece A1
  Simulation: attach piece A2
  Simulation: attach piece A3
  Simulation: attach piece A4
  Simulation: attach piece A5
  Simulation: attach piece A6
  Simulation: attach piece B1
  Simulation: attach piece B2
  Simulation: attach piece B3
  Simulation: attach piece B4
  Simulation: attach piece B5
  Simulation: attach piece B6
  MoveL (bench lift)
  Set speed (100.0 mm/s)
  MoveL (bench over AMR)
  Set speed (20.0 mm/s)
  MoveL (bench down)
  Set IO_0=0
  Pause 500 ms
  Simulation: release bench
  MoveL (bench place out)
  Set speed (100.0 mm/s)
  MoveL (bench place out up)
  MoveL (back to middle)
  MoveJ (Home)

--- Python program Deliver (AMR) ---
"""The AMR drives the finished bench 2 m away along the table and comes back (RoboDK station script
"Deliver (AMR)").

    python robot_cell/amr_drive.py           also works from outside RoboDK

Needs only the robodk package. Everything under the station's "AMR" frame rides along: its plate,
top module and LD-250, and the bench once the robot program has set it down there (the program's
release puts the bench under the AMR frame).
"""
import time

from robodk import robolink, robomath

DISTANCE = 2000          # mm, along the ground base's x (away from the robot)
STEPS = 120              # per direction
PAUSE = 1.0              # s at the far end
OWN = ("AMR plate", "AMR top module")


def main():
    RDK = robolink.Robolink()
    amr = RDK.Item("AMR", robolink.ITEM_TYPE_FRAME)
    if not amr.Valid():
        raise SystemExit("no AMR in the open station")
    riding = [c for c in amr.Childs() if c.Type() == robolink.ITEM_TYPE_OBJECT and c.Name() not in OWN]
    home = amr.Pose()
    for out in (True, False):
        for i in range(1, STEPS + 1):
            s = i / STEPS if out else 1 - i / STEPS
            s = 0.5 - 0.5 * robomath.cos(robomath.pi * s)        # smooth start and stop
            amr.setPose(robomath.transl(DISTANCE * s, 0, 0) * home)
            RDK.Render(True)
            time.sleep(0.02)
        if out:
            time.sleep(PAUSE)
    amr.setPose(home)
    print(f"AMR drove {DISTANCE / 1000:.0f} m and back with {len(riding)} parts on its plate")


if __name__ == "__main__":
    main()

--- Python program Assemble and deliver ---
"""The whole cycle (station script "Assemble and deliver"): the robot program AssembleBench builds the
bench and sets it down on the AMR, then the AMR drives it 2 m along the table and back (amr_drive.py).

    python robot_cell/assemble_and_deliver.py      also works from outside RoboDK
"""
import time

from robodk import robolink

import amr_drive


def main():
    RDK = robolink.Robolink()
    prog = RDK.Item("AssembleBench", robolink.ITEM_TYPE_PROGRAM)
    if not prog.Valid():
        raise SystemExit("no AssembleBench in the open station")
    t0 = time.time()
    prog.RunProgram()
    time.sleep(1)
    while prog.Busy():
        time.sleep(0.2)
    print(f"AssembleBench done after {time.time() - t0:.0f} s (at the simulation speed)")
    amr_drive.main()


if __name__ == "__main__":
    main()
